Staubli VAL3: actionItem.pjx

--- actionItem.pjx ---
Parameters version=s8.10.3Cs9_BS2093 stackSize=5000 millimeterUnit=true
Data file=actionItem.dtx

--- actionItem.dtx ---
public num nIOindex
public num nboolValue
public num nPulseValue
public string sIOtype
public string sValue
public bool bActive
